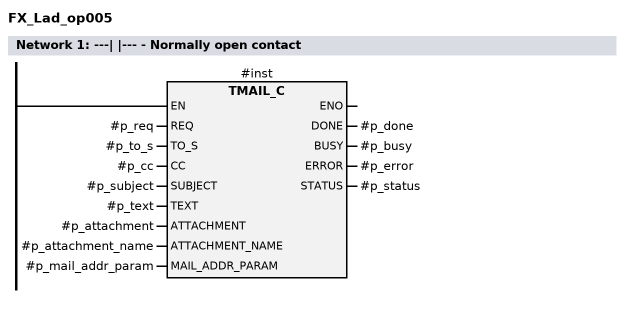
   #inst(REQ := #p_req,   // TMAIL_C
         TO_S := #p_to_s,
         CC := #p_cc,
         SUBJECT := #p_subject,
         TEXT := #p_text,
         ATTACHMENT := #p_attachment,
         ATTACHMENT_NAME := #p_attachment_name,
         MAIL_ADDR_PARAM := #p_mail_addr_param,
         DONE => #p_done,
         BUSY => #p_busy,
         ERROR => #p_error,
         STATUS => #p_status);
END_REGION
END_FUNCTION_BLOCK

FUNCTION_BLOCK "FX_Lad_op021"   // FB349, LAD
{ S7_Optimized_Access := 'TRUE' }
VERSION : 0.1
   VAR_INPUT
      "a" : Bool;
      "b" : Bool;
      c : Bool;
      ia : Int;
      ib : Int;
      ic : Int;
      da : DInt;
      db : DInt;
      ra : Real;
      rb : Real;
      wa : Word;
      wb : Word;
      dwa : DWord;
      ba : Byte;
      ta : Time;
      tb : Time;
      s1 : String;
      s2 : String;
   END_VAR
   VAR_OUTPUT
      q : Bool;
      q2 : Bool;
      io : Int;
      io2 : Int;
      dout : DInt;
      rout : Real;
      wout : Word;
      dwout : DWord;
      bout : Byte;
      tout : Time;
      sout : String;
   END_VAR
   VAR_IN_OUT
      p_req : Bool;
      p_interface : Hw_Interface;
      p_conf_data : Variant;
      p_done : Bool;
      p_busy : Bool;
      p_error : Bool;
      p_status : DWord;
      p_err_loc : DWord;
      arr : Array[0..9] of Int;
      barr : Array[0..7] of Bool;
      iinout : Int;
   END_VAR
   VAR
      inst : T_CONFIG;
      ton1 : TON_TIME;
      tof1 : TOF_TIME;
      tp1 : TP_TIME;
      tonr1 : TONR_TIME;
      ctu1 : CTU_INT;
      ctd1 : CTD_INT;
      ctud1 : CTUD_INT;
      rtrig1 : R_TRIG;
      ftrig1 : F_TRIG;
      edge1 : Bool;
      edge2 : Bool;
      stat1 : Bool;
      stat2 : Bool;
      stati : Int;
   END_VAR
   VAR_TEMP
      t1 : Bool;
      t2 : Bool;
      ti : Int;
      td : DInt;
      tr : Real;
      tw : Word;
      tt : Time;
      var1 : Variant;
   END_VAR
BEGIN

REGION Network 1: ---| |--- - Normally open contact
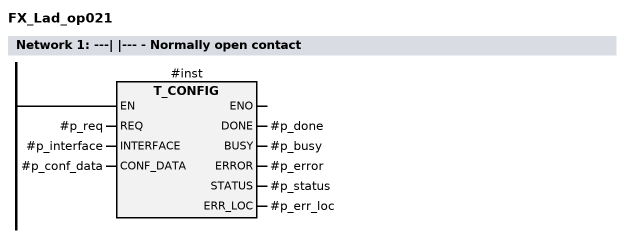
   #inst(Req := #p_req,   // T_CONFIG
         Interface := #p_interface,
         Conf_Data := #p_conf_data,
         Done => #p_done,
         Busy => #p_busy,
         Error => #p_error,
         Status => #p_status,
         Err_Loc => #p_err_loc);
END_REGION
END_FUNCTION_BLOCK

FUNCTION_BLOCK "FB_Lad_Trcv"   // FB350, LAD
{ S7_Optimized_Access := 'TRUE' }
   VAR_INPUT
      en_r : Bool;
      cont : Bool;
      len : UInt;
      id : Conn_Ouc;
      adhoc : Bool;
   END_VAR
   VAR_OUTPUT
      done : Bool;
      busy : Bool;
      err : Bool;
      status : Word;
      rcvdlen : UInt;
   END_VAR
   VAR_IN_OUT
      connect : TCON_IP_v4;
      data : Array[0..99] of Byte;
      comrst : Bool;
      addr : Variant;
   END_VAR
   VAR
      inst : TRCV;
   END_VAR
BEGIN

REGION Network 1: TRCV
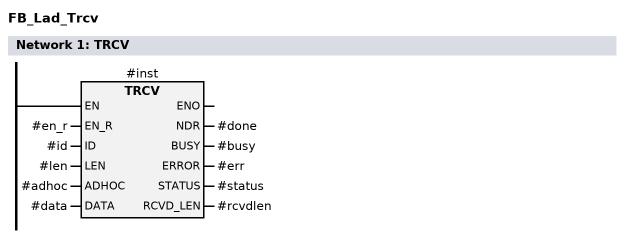
   #inst(EN_R := #en_r,   // TRCV
         ID := #id,
         LEN := #len,
         ADHOC := #adhoc,
         DATA := #data,
         NDR => #done,
         BUSY => #busy,
         ERROR => #err,
         STATUS => #status,
         RCVD_LEN => #rcvdlen);
END_REGION
END_FUNCTION_BLOCK

FUNCTION_BLOCK "FB_Lad_TrcvC"   // FB351, LAD
{ S7_Optimized_Access := 'TRUE' }
   VAR_INPUT
      en_r : Bool;
      cont : Bool;
      len : UInt;
      id : Conn_Ouc;
      adhoc : Bool;
   END_VAR
   VAR_OUTPUT
      done : Bool;
      busy : Bool;
      err : Bool;
      status : Word;
      rcvdlen : UInt;
   END_VAR
   VAR_IN_OUT
      connect : TCON_IP_v4;
      data : Array[0..99] of Byte;
      comrst : Bool;
      addr : Variant;
   END_VAR
   VAR
      inst : TRCV_C;
   END_VAR
BEGIN

REGION Network 1: TRCV_C
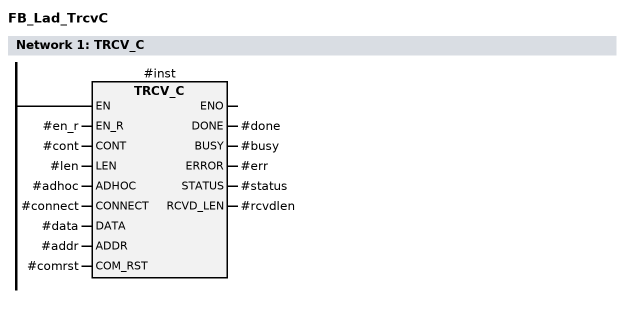
   #inst(EN_R := #en_r,   // TRCV_C
         CONT := #cont,
         LEN := #len,
         ADHOC := #adhoc,
         CONNECT := #connect,
         DATA := #data,
         ADDR := #addr,
         COM_RST := #comrst,
         DONE => #done,
         BUSY => #busy,
         ERROR => #err,
         STATUS => #status,
         RCVD_LEN => #rcvdlen);
END_REGION
END_FUNCTION_BLOCK

FUNCTION_BLOCK "FB_Fbd_TrcvC"   // FB352, FBD
{ S7_Optimized_Access := 'TRUE' }
   VAR_INPUT
      en_r : Bool;
      cont : Bool;
      len : UInt;
      id : Conn_Ouc;
      adhoc : Bool;
   END_VAR
   VAR_OUTPUT
      done : Bool;
      busy : Bool;
      err : Bool;
      status : Word;
      rcvdlen : UInt;
   END_VAR
   VAR_IN_OUT
      connect : TCON_IP_v4;
      data : Array[0..99] of Byte;
      comrst : Bool;
      addr : Variant;
   END_VAR
   VAR
      inst : TRCV_C;
   END_VAR
BEGIN

REGION Network 1: TRCV_C
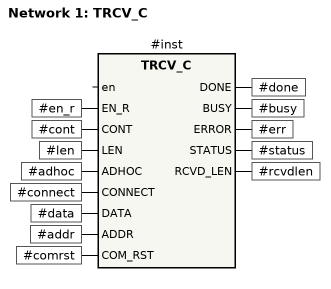
   #inst(EN_R := #en_r,   // TRCV_C
         CONT := #cont,
         LEN := #len,
         ADHOC := #adhoc,
         CONNECT := #connect,
         DATA := #data,
         ADDR := #addr,
         COM_RST := #comrst,
         DONE => #done,
         BUSY => #busy,
         ERROR => #err,
         STATUS => #status,
         RCVD_LEN => #rcvdlen);
END_REGION
END_FUNCTION_BLOCK

FUNCTION_BLOCK "FB_Fbd_Trcv"   // FB353, FBD
{ S7_Optimized_Access := 'TRUE' }
   VAR_INPUT
      en_r : Bool;
      cont : Bool;
      len : UInt;
      id : Conn_Ouc;
      adhoc : Bool;
   END_VAR
   VAR_OUTPUT
      done : Bool;
      busy : Bool;
      err : Bool;
      status : Word;
      rcvdlen : UInt;
   END_VAR
   VAR_IN_OUT
      connect : TCON_IP_v4;
      data : Array[0..99] of Byte;
      comrst : Bool;
      addr : Variant;
   END_VAR
   VAR
      inst : TRCV;
   END_VAR
BEGIN

REGION Network 1: TRCV
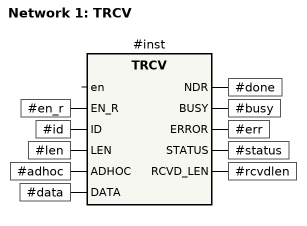
   #inst(EN_R := #en_r,   // TRCV
         ID := #id,
         LEN := #len,
         ADHOC := #adhoc,
         DATA := #data,
         NDR => #done,
         BUSY => #busy,
         ERROR => #err,
         STATUS => #status,
         RCVD_LEN => #rcvdlen);
END_REGION
END_FUNCTION_BLOCK

FUNCTION_BLOCK "FX_Fbd_op005"   // FB354, FBD
{ S7_Optimized_Access := 'TRUE' }
VERSION : 0.1
   VAR_INPUT
      "a" : Bool;
      "b" : Bool;
      c : Bool;
      ia : Int;
      ib : Int;
      ic : Int;
      da : DInt;
      db : DInt;
      ra : Real;
      rb : Real;
      wa : Word;
      wb : Word;
      dwa : DWord;
      ba : Byte;
      ta : Time;
      tb : Time;
      s1 : String;
      s2 : String;
   END_VAR
   VAR_OUTPUT
      q : Bool;
      q2 : Bool;
      io : Int;
      io2 : Int;
      dout : DInt;
      rout : Real;
      wout : Word;
      dwout : DWord;
      bout : Byte;
      tout : Time;
      sout : String;
   END_VAR
   VAR_IN_OUT
      p_req : Bool;
      p_to_s : String;
      p_cc : String;
      p_subject : String;
      p_text : String;
      p_attachment : Variant;
      p_attachment_name : String;
      p_mail_addr_param : Variant;
      p_done : Bool;
      p_busy : Bool;
      p_error : Bool;
      p_status : Word;
      arr : Array[0..9] of Int;
      barr : Array[0..7] of Bool;
      iinout : Int;
   END_VAR
   VAR
      inst : TMAIL_C;
      ton1 : TON_TIME;
      tof1 : TOF_TIME;
      tp1 : TP_TIME;
      tonr1 : TONR_TIME;
      ctu1 : CTU_INT;
      ctd1 : CTD_INT;
      ctud1 : CTUD_INT;
      rtrig1 : R_TRIG;
      ftrig1 : F_TRIG;
      edge1 : Bool;
      edge2 : Bool;
      stat1 : Bool;
      stat2 : Bool;
      stati : Int;
   END_VAR
   VAR_TEMP
      t1 : Bool;
      t2 : Bool;
      ti : Int;
      td : DInt;
      tr : Real;
      tw : Word;
      tt : Time;
      var1 : Variant;
   END_VAR
BEGIN

REGION Network 1: ---| |--- - Normally open contact
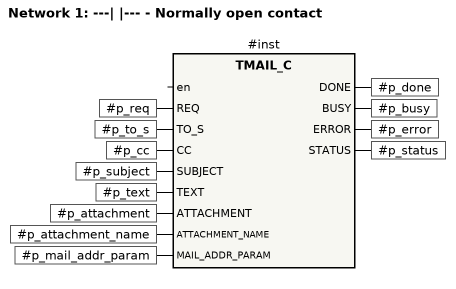
   #inst(REQ := #p_req,   // TMAIL_C
         TO_S := #p_to_s,
         CC := #p_cc,
         SUBJECT := #p_subject,
         TEXT := #p_text,
         ATTACHMENT := #p_attachment,
         ATTACHMENT_NAME := #p_attachment_name,
         MAIL_ADDR_PARAM := #p_mail_addr_param,
         DONE => #p_done,
         BUSY => #p_busy,
         ERROR => #p_error,
         STATUS => #p_status);
END_REGION
END_FUNCTION_BLOCK

FUNCTION_BLOCK "FX_Fbd_op021"   // FB355, FBD
{ S7_Optimized_Access := 'TRUE' }
VERSION : 0.1
   VAR_INPUT
      "a" : Bool;
      "b" : Bool;
      c : Bool;
      ia : Int;
      ib : Int;
      ic : Int;
      da : DInt;
      db : DInt;
      ra : Real;
      rb : Real;
      wa : Word;
      wb : Word;
      dwa : DWord;
      ba : Byte;
      ta : Time;
      tb : Time;
      s1 : String;
      s2 : String;
   END_VAR
   VAR_OUTPUT
      q : Bool;
      q2 : Bool;
      io : Int;
      io2 : Int;
      dout : DInt;
      rout : Real;
      wout : Word;
      dwout : DWord;
      bout : Byte;
      tout : Time;
      sout : String;
   END_VAR
   VAR_IN_OUT
      p_req : Bool;
      p_interface : Hw_Interface;
      p_conf_data : Variant;
      p_done : Bool;
      p_busy : Bool;
      p_error : Bool;
      p_status : DWord;
      p_err_loc : DWord;
      arr : Array[0..9] of Int;
      barr : Array[0..7] of Bool;
      iinout : Int;
   END_VAR
   VAR
      inst : T_CONFIG;
      ton1 : TON_TIME;
      tof1 : TOF_TIME;
      tp1 : TP_TIME;
      tonr1 : TONR_TIME;
      ctu1 : CTU_INT;
      ctd1 : CTD_INT;
      ctud1 : CTUD_INT;
      rtrig1 : R_TRIG;
      ftrig1 : F_TRIG;
      edge1 : Bool;
      edge2 : Bool;
      stat1 : Bool;
      stat2 : Bool;
      stati : Int;
   END_VAR
   VAR_TEMP
      t1 : Bool;
      t2 : Bool;
      ti : Int;
      td : DInt;
      tr : Real;
      tw : Word;
      tt : Time;
      var1 : Variant;
   END_VAR
BEGIN

REGION Network 1: ---| |--- - Normally open contact
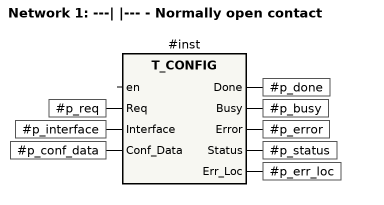
   #inst(Req := #p_req,   // T_CONFIG
         Interface := #p_interface,
         Conf_Data := #p_conf_data,
         Done => #p_done,
         Busy => #p_busy,
         Error => #p_error,
         Status => #p_status,
         Err_Loc => #p_err_loc);
END_REGION
END_FUNCTION_BLOCK

FUNCTION_BLOCK "FB_Lad_ex051"   // FB356, LAD
{ S7_Optimized_Access := 'TRUE' }
   VAR_INPUT
      v_mode : Int;
      v_f_id : Hw_Io;
      v_mlen : UInt;
   END_VAR
   VAR_OUTPUT
      v_new : Bool;
      v_status : DWord;
      v_id : Hw_Io;
      v_len : UInt;
   END_VAR
   VAR_IN_OUT
      v_tinfo : Array[0..99] of Byte;
      v_ainfo : Array[0..99] of Byte;
   END_VAR
   VAR
      inst : RALRM;
   END_VAR
BEGIN

REGION Network 1: Description RALRM
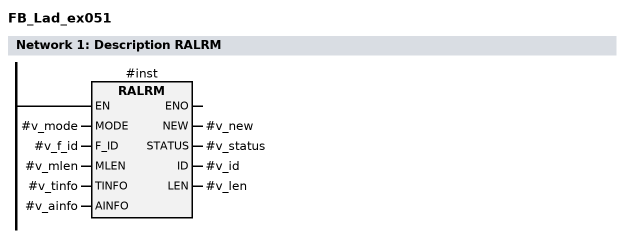
   #inst(MODE := #v_mode,   // RALRM
         F_ID := #v_f_id,
         MLEN := #v_mlen,
         TINFO := #v_tinfo,
         AINFO := #v_ainfo,
         NEW => #v_new,
         STATUS => #v_status,
         ID => #v_id,
         LEN => #v_len);
END_REGION
END_FUNCTION_BLOCK

FUNCTION_BLOCK "FB_Lad_ex071"   // FB357, LAD
{ S7_Optimized_Access := 'TRUE' }
   VAR_INPUT
      v_com_rst : Bool;
      v_start : Bool;
      v_end : Bool;
   END_VAR
   VAR_OUTPUT
      v_status : DWord;
   END_VAR
   VAR_IN_OUT
      v_penergy : PE_PLUS;
   END_VAR
   VAR
      inst : PE_WOL;
   END_VAR
BEGIN

REGION Network 1: Description PE_WOL
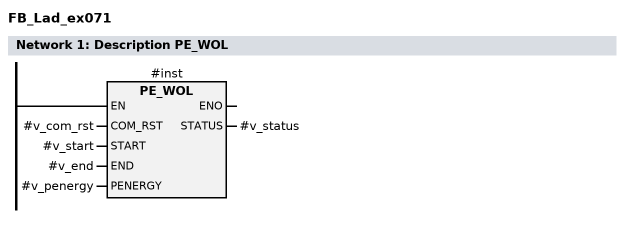
   #inst(COM_RST := #v_com_rst, START := #v_start, END := #v_end, PENERGY := #v_penergy, STATUS => #v_status);   // PE_WOL
END_REGION
END_FUNCTION_BLOCK

FUNCTION_BLOCK "FX_Lad_ex037"   // FB358, LAD
{ S7_Optimized_Access := 'TRUE' }
VERSION : 0.1
   VAR_INPUT
      "a" : Bool;
      "b" : Bool;
      c : Bool;
      ia : Int;
      ib : Int;
      ic : Int;
      da : DInt;
      db : DInt;
      ra : Real;
      rb : Real;
      wa : Word;
      wb : Word;
      dwa : DWord;
      ba : Byte;
      ta : Time;
      tb : Time;
      s1 : String;
      s2 : String;
   END_VAR
   VAR_OUTPUT
      q : Bool;
      q2 : Bool;
      io : Int;
      io2 : Int;
      dout : DInt;
      rout : Real;
      wout : Word;
      dwout : DWord;
      bout : Byte;
      tout : Time;
      sout : String;
   END_VAR
   VAR_IN_OUT
      x_wstring : WString;
      arr : Array[0..9] of Int;
      barr : Array[0..7] of Bool;
      iinout : Int;
   END_VAR
   VAR
      ton1 : TON_TIME;
      tof1 : TOF_TIME;
      tp1 : TP_TIME;
      tonr1 : TONR_TIME;
      ctu1 : CTU_INT;
      ctd1 : CTD_INT;
      ctud1 : CTUD_INT;
      rtrig1 : R_TRIG;
      ftrig1 : F_TRIG;
      edge1 : Bool;
      edge2 : Bool;
      stat1 : Bool;
      stat2 : Bool;
      stati : Int;
   END_VAR
   VAR_TEMP
      t1 : Bool;
      t2 : Bool;
      ti : Int;
      td : DInt;
      tr : Real;
      tw : Word;
      tt : Time;
      var1 : Variant;
   END_VAR
BEGIN

REGION Network 1: ---| |--- - Normally open contact
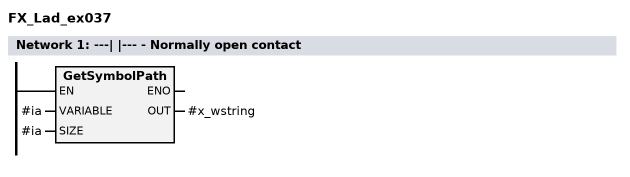
   // no SCL statement known for GetSymbolPath: written as a call
   #x_wstring := GetSymbolPath(variable := #ia, size := #ia);
END_REGION
END_FUNCTION_BLOCK

FUNCTION_BLOCK "FX_Lad_ex051"   // FB359, LAD
{ S7_Optimized_Access := 'TRUE' }
VERSION : 0.1
   VAR_INPUT
      "a" : Bool;
      "b" : Bool;
      c : Bool;
      ia : Int;
      ib : Int;
      ic : Int;
      da : DInt;
      db : DInt;
      ra : Real;
      rb : Real;
      wa : Word;
      wb : Word;
      dwa : DWord;
      ba : Byte;
      ta : Time;
      tb : Time;
      s1 : String;
      s2 : String;
   END_VAR
   VAR_OUTPUT
      q : Bool;
      q2 : Bool;
      io : Int;
      io2 : Int;
      dout : DInt;
      rout : Real;
      wout : Word;
      dwout : DWord;
      bout : Byte;
      tout : Time;
      sout : String;
   END_VAR
   VAR_IN_OUT
      p_mode : Int;
      p_f_id : Hw_Io;
      p_mlen : UInt;
      p_new : Bool;
      p_status : DWord;
      p_id : Hw_Io;
      p_len : UInt;
      p_tinfo : Variant;
      p_ainfo : Variant;
      arr : Array[0..9] of Int;
      barr : Array[0..7] of Bool;
      iinout : Int;
   END_VAR
   VAR
      inst : RALRM;
      ton1 : TON_TIME;
      tof1 : TOF_TIME;
      tp1 : TP_TIME;
      tonr1 : TONR_TIME;
      ctu1 : CTU_INT;
      ctd1 : CTD_INT;
      ctud1 : CTUD_INT;
      rtrig1 : R_TRIG;
      ftrig1 : F_TRIG;
      edge1 : Bool;
      edge2 : Bool;
      stat1 : Bool;
      stat2 : Bool;
      stati : Int;
   END_VAR
   VAR_TEMP
      t1 : Bool;
      t2 : Bool;
      ti : Int;
      td : DInt;
      tr : Real;
      tw : Word;
      tt : Time;
      var1 : Variant;
   END_VAR
BEGIN

REGION Network 1: ---| |--- - Normally open contact
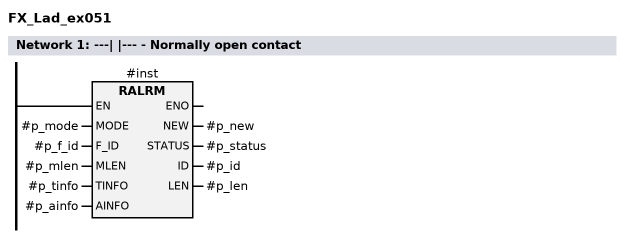
   #inst(MODE := #p_mode,   // RALRM
         F_ID := #p_f_id,
         MLEN := #p_mlen,
         TINFO := #p_tinfo,
         AINFO := #p_ainfo,
         NEW => #p_new,
         STATUS => #p_status,
         ID => #p_id,
         LEN => #p_len);
END_REGION
END_FUNCTION_BLOCK

FUNCTION_BLOCK "FB_Fbd_ex037"   // FB360, FBD
{ S7_Optimized_Access := 'TRUE' }
   VAR_INPUT
      v_size : DInt;
   END_VAR
   VAR_OUTPUT
      v_out : WString;
   END_VAR
   VAR_IN_OUT
      v_variable : Variant;
   END_VAR
BEGIN

REGION Network 1: Querying GetSymbolPath - actual parameter at beginning of a call path
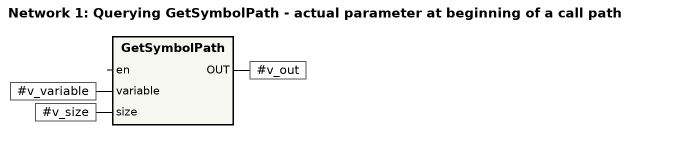
   // no SCL statement known for GetSymbolPath: written as a call
   #v_out := GetSymbolPath(variable := #v_variable, size := #v_size);
END_REGION
END_FUNCTION_BLOCK

FUNCTION_BLOCK "FB_Fbd_ex051"   // FB361, FBD
{ S7_Optimized_Access := 'TRUE' }
   VAR_INPUT
      v_mode : Int;
      v_f_id : Hw_Io;
      v_mlen : UInt;
   END_VAR
   VAR_OUTPUT
      v_new : Bool;
      v_status : DWord;
      v_id : Hw_Io;
      v_len : UInt;
   END_VAR
   VAR_IN_OUT
      v_tinfo : Array[0..99] of Byte;
      v_ainfo : Array[0..99] of Byte;
   END_VAR
   VAR
      inst : RALRM;
   END_VAR
BEGIN

REGION Network 1: Description RALRM
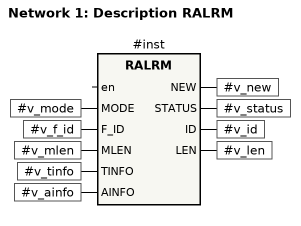
   #inst(MODE := #v_mode,   // RALRM
         F_ID := #v_f_id,
         MLEN := #v_mlen,
         TINFO := #v_tinfo,
         AINFO := #v_ainfo,
         NEW => #v_new,
         STATUS => #v_status,
         ID => #v_id,
         LEN => #v_len);
END_REGION
END_FUNCTION_BLOCK

FUNCTION_BLOCK "FB_Fbd_ex071"   // FB362, FBD
{ S7_Optimized_Access := 'TRUE' }
   VAR_INPUT
      v_com_rst : Bool;
      v_start : Bool;
      v_end : Bool;
   END_VAR
   VAR_OUTPUT
      v_status : DWord;
   END_VAR
   VAR_IN_OUT
      v_penergy : PE_PLUS;
   END_VAR
   VAR
      inst : PE_WOL;
   END_VAR
BEGIN

REGION Network 1: Description PE_WOL
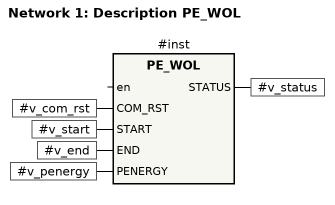
   #inst(COM_RST := #v_com_rst, START := #v_start, END := #v_end, PENERGY := #v_penergy, STATUS => #v_status);   // PE_WOL
END_REGION
END_FUNCTION_BLOCK

FUNCTION_BLOCK "FX_Lad_095"   // FB363, LAD
{ S7_Optimized_Access := 'TRUE' }
VERSION : 0.1
   VAR_INPUT
      "a" : Bool;
      "b" : Bool;
      c : Bool;
      ia : Int;
      ib : Int;
      ic : Int;
      da : DInt;
      db : DInt;
      ra : Real;
      rb : Real;
      wa : Word;
      wb : Word;
      dwa : DWord;
      ba : Byte;
      ta : Time;
      tb : Time;
      s1 : String;
      s2 : String;
   END_VAR
   VAR_OUTPUT
      q : Bool;
      q2 : Bool;
      io : Int;
      io2 : Int;
      dout : DInt;
      rout : Real;
      wout : Word;
      dwout : DWord;
      bout : Byte;
      tout : Time;
      sout : String;
   END_VAR
   VAR_IN_OUT
      x_usint : USInt;
      arr : Array[0..9] of Int;
      barr : Array[0..7] of Bool;
      iinout : Int;
   END_VAR
   VAR
      ton1 : TON_TIME;
      tof1 : TOF_TIME;
      tp1 : TP_TIME;
      tonr1 : TONR_TIME;
      ctu1 : CTU_INT;
      ctd1 : CTD_INT;
      ctud1 : CTUD_INT;
      rtrig1 : R_TRIG;
      ftrig1 : F_TRIG;
      edge1 : Bool;
      edge2 : Bool;
      stat1 : Bool;
      stat2 : Bool;
      stati : Int;
   END_VAR
   VAR_TEMP
      t1 : Bool;
      t2 : Bool;
      ti : Int;
      td : DInt;
      tr : Real;
      tw : Word;
      tt : Time;
      var1 : Variant;
   END_VAR
BEGIN

REGION Network 1: ---| |--- - Normally open contact
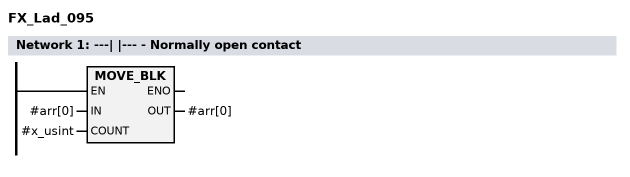
   MOVE_BLK(IN := #arr[0], COUNT := #x_usint, OUT => #arr[0]);
END_REGION
END_FUNCTION_BLOCK

FUNCTION_BLOCK "FX_Lad_097"   // FB364, LAD
{ S7_Optimized_Access := 'TRUE' }
VERSION : 0.1
   VAR_INPUT
      "a" : Bool;
      "b" : Bool;
      c : Bool;
      ia : Int;
      ib : Int;
      ic : Int;
      da : DInt;
      db : DInt;
      ra : Real;
      rb : Real;
      wa : Word;
      wb : Word;
      dwa : DWord;
      ba : Byte;
      ta : Time;
      tb : Time;
      s1 : String;
      s2 : String;
   END_VAR
   VAR_OUTPUT
      q : Bool;
      q2 : Bool;
      io : Int;
      io2 : Int;
      dout : DInt;
      rout : Real;
      wout : Word;
      dwout : DWord;
      bout : Byte;
      tout : Time;
      sout : String;
   END_VAR
   VAR_IN_OUT
      x_usint : USInt;
      arr : Array[0..9] of Int;
      barr : Array[0..7] of Bool;
      iinout : Int;
   END_VAR
   VAR
      ton1 : TON_TIME;
      tof1 : TOF_TIME;
      tp1 : TP_TIME;
      tonr1 : TONR_TIME;
      ctu1 : CTU_INT;
      ctd1 : CTD_INT;
      ctud1 : CTUD_INT;
      rtrig1 : R_TRIG;
      ftrig1 : F_TRIG;
      edge1 : Bool;
      edge2 : Bool;
      stat1 : Bool;
      stat2 : Bool;
      stati : Int;
   END_VAR
   VAR_TEMP
      t1 : Bool;
      t2 : Bool;
      ti : Int;
      td : DInt;
      tr : Real;
      tw : Word;
      tt : Time;
      var1 : Variant;
   END_VAR
BEGIN

REGION Network 1: ---| |--- - Normally open contact
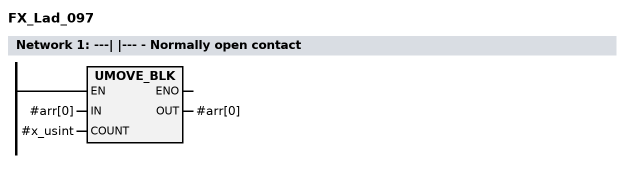
   UMOVE_BLK(IN := #arr[0], COUNT := #x_usint, OUT => #arr[0]);
END_REGION
END_FUNCTION_BLOCK

FUNCTION_BLOCK "FX_Lad_098"   // FB365, LAD
{ S7_Optimized_Access := 'TRUE' }
VERSION : 0.1
   VAR_INPUT
      "a" : Bool;
      "b" : Bool;
      c : Bool;
      ia : Int;
      ib : Int;
      ic : Int;
      da : DInt;
      db : DInt;
      ra : Real;
      rb : Real;
      wa : Word;
      wb : Word;
      dwa : DWord;
      ba : Byte;
      ta : Time;
      tb : Time;
      s1 : String;
      s2 : String;
   END_VAR
   VAR_OUTPUT
      q : Bool;
      q2 : Bool;
      io : Int;
      io2 : Int;
      dout : DInt;
      rout : Real;
      wout : Word;
      dwout : DWord;
      bout : Byte;
      tout : Time;
      sout : String;
   END_VAR
   VAR_IN_OUT
      p_in : Date;
      p_count : USInt;
      p_out : Date;
      s_in : Int;
      s_count : UDInt;
      s_out : Array[0..9] of Int;
      arr : Array[0..9] of Int;
      barr : Array[0..7] of Bool;
      iinout : Int;
   END_VAR
   VAR
      ton1 : TON_TIME;
      tof1 : TOF_TIME;
      tp1 : TP_TIME;
      tonr1 : TONR_TIME;
      ctu1 : CTU_INT;
      ctd1 : CTD_INT;
      ctud1 : CTUD_INT;
      rtrig1 : R_TRIG;
      ftrig1 : F_TRIG;
      edge1 : Bool;
      edge2 : Bool;
      stat1 : Bool;
      stat2 : Bool;
      stati : Int;
   END_VAR
   VAR_TEMP
      t1 : Bool;
      t2 : Bool;
      ti : Int;
      td : DInt;
      tr : Real;
      tw : Word;
      tt : Time;
      var1 : Variant;
   END_VAR
BEGIN

REGION Network 1: ---| |--- - Normally open contact
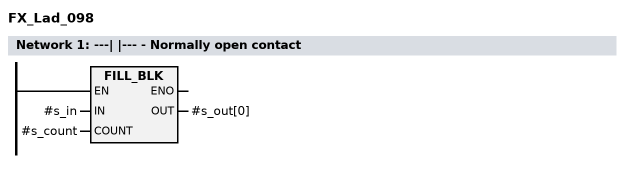
   RUNG wire#powerrail
      FillBlockI(in := #s_in, count := #s_count, out => #s_out[0])
   END_RUNG
   // the same network as SCL:
   FILL_BLK(IN := #s_in, COUNT := #s_count, OUT => #s_out[0]);
END_REGION
END_FUNCTION_BLOCK

FUNCTION_BLOCK "FX_Lad_099"   // FB366, LAD
{ S7_Optimized_Access := 'TRUE' }
VERSION : 0.1
   VAR_INPUT
      "a" : Bool;
      "b" : Bool;
      c : Bool;
      ia : Int;
      ib : Int;
      ic : Int;
      da : DInt;
      db : DInt;
      ra : Real;
      rb : Real;
      wa : Word;
      wb : Word;
      dwa : DWord;
      ba : Byte;
      ta : Time;
      tb : Time;
      s1 : String;
      s2 : String;
   END_VAR
   VAR_OUTPUT
      q : Bool;
      q2 : Bool;
      io : Int;
      io2 : Int;
      dout : DInt;
      rout : Real;
      wout : Word;
      dwout : DWord;
      bout : Byte;
      tout : Time;
      sout : String;
   END_VAR
   VAR_IN_OUT
      p_in : Date;
      p_count : USInt;
      p_out : Date;
      s_in : Int;
      s_count : UDInt;
      s_out : Array[0..9] of Int;
      arr : Array[0..9] of Int;
      barr : Array[0..7] of Bool;
      iinout : Int;
   END_VAR
   VAR
      ton1 : TON_TIME;
      tof1 : TOF_TIME;
      tp1 : TP_TIME;
      tonr1 : TONR_TIME;
      ctu1 : CTU_INT;
      ctd1 : CTD_INT;
      ctud1 : CTUD_INT;
      rtrig1 : R_TRIG;
      ftrig1 : F_TRIG;
      edge1 : Bool;
      edge2 : Bool;
      stat1 : Bool;
      stat2 : Bool;
      stati : Int;
   END_VAR
   VAR_TEMP
      t1 : Bool;
      t2 : Bool;
      ti : Int;
      td : DInt;
      tr : Real;
      tw : Word;
      tt : Time;
      var1 : Variant;
   END_VAR
BEGIN

REGION Network 1: ---| |--- - Normally open contact
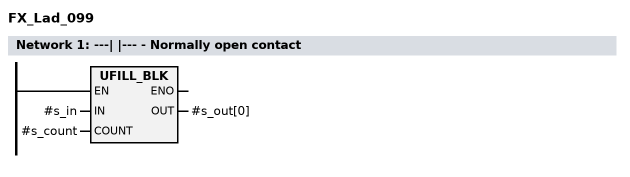
   UFILL_BLK(IN := #s_in, COUNT := #s_count, OUT => #s_out[0]);
END_REGION
END_FUNCTION_BLOCK

FUNCTION_BLOCK "FX_Fbd_100"   // FB367, FBD
{ S7_Optimized_Access := 'TRUE' }
VERSION : 0.1
   VAR_INPUT
      "a" : Bool;
      "b" : Bool;
      c : Bool;
      ia : Int;
      ib : Int;
      ic : Int;
      da : DInt;
      db : DInt;
      ra : Real;
      rb : Real;
      wa : Word;
      wb : Word;
      dwa : DWord;
      ba : Byte;
      ta : Time;
      tb : Time;
      s1 : String;
      s2 : String;
   END_VAR
   VAR_OUTPUT
      q : Bool;
      q2 : Bool;
      io : Int;
      io2 : Int;
      dout : DInt;
      rout : Real;
      wout : Word;
      dwout : DWord;
      bout : Byte;
      tout : Time;
      sout : String;
   END_VAR
   VAR_IN_OUT
      x_usint : USInt;
      arr : Array[0..9] of Int;
      barr : Array[0..7] of Bool;
      iinout : Int;
   END_VAR
   VAR
      ton1 : TON_TIME;
      tof1 : TOF_TIME;
      tp1 : TP_TIME;
      tonr1 : TONR_TIME;
      ctu1 : CTU_INT;
      ctd1 : CTD_INT;
      ctud1 : CTUD_INT;
      rtrig1 : R_TRIG;
      ftrig1 : F_TRIG;
      edge1 : Bool;
      edge2 : Bool;
      stat1 : Bool;
      stat2 : Bool;
      stati : Int;
   END_VAR
   VAR_TEMP
      t1 : Bool;
      t2 : Bool;
      ti : Int;
      td : DInt;
      tr : Real;
      tw : Word;
      tt : Time;
      var1 : Variant;
   END_VAR
BEGIN

REGION Network 1: ---| |--- - Normally open contact
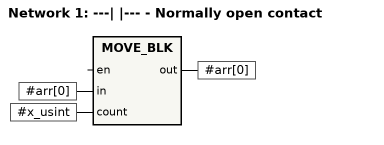
   MOVE_BLK(IN := #arr[0], COUNT := #x_usint, OUT => #arr[0]);
END_REGION
END_FUNCTION_BLOCK

FUNCTION_BLOCK "FX_Fbd_102"   // FB368, FBD
{ S7_Optimized_Access := 'TRUE' }
VERSION : 0.1
   VAR_INPUT
      "a" : Bool;
      "b" : Bool;
      c : Bool;
      ia : Int;
      ib : Int;
      ic : Int;
      da : DInt;
      db : DInt;
      ra : Real;
      rb : Real;
      wa : Word;
      wb : Word;
      dwa : DWord;
      ba : Byte;
      ta : Time;
      tb : Time;
      s1 : String;
      s2 : String;
   END_VAR
   VAR_OUTPUT
      q : Bool;
      q2 : Bool;
      io : Int;
      io2 : Int;
      dout : DInt;
      rout : Real;
      wout : Word;
      dwout : DWord;
      bout : Byte;
      tout : Time;
      sout : String;
   END_VAR
   VAR_IN_OUT
      x_usint : USInt;
      arr : Array[0..9] of Int;
      barr : Array[0..7] of Bool;
      iinout : Int;
   END_VAR
   VAR
      ton1 : TON_TIME;
      tof1 : TOF_TIME;
      tp1 : TP_TIME;
      tonr1 : TONR_TIME;
      ctu1 : CTU_INT;
      ctd1 : CTD_INT;
      ctud1 : CTUD_INT;
      rtrig1 : R_TRIG;
      ftrig1 : F_TRIG;
      edge1 : Bool;
      edge2 : Bool;
      stat1 : Bool;
      stat2 : Bool;
      stati : Int;
   END_VAR
   VAR_TEMP
      t1 : Bool;
      t2 : Bool;
      ti : Int;
      td : DInt;
      tr : Real;
      tw : Word;
      tt : Time;
      var1 : Variant;
   END_VAR
BEGIN

REGION Network 1: ---| |--- - Normally open contact
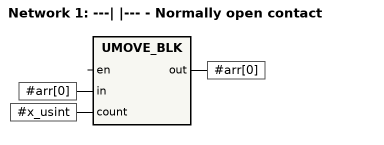
   UMOVE_BLK(IN := #arr[0], COUNT := #x_usint, OUT => #arr[0]);
END_REGION
END_FUNCTION_BLOCK

FUNCTION_BLOCK "FX_Fbd_103"   // FB369, FBD
{ S7_Optimized_Access := 'TRUE' }
VERSION : 0.1
   VAR_INPUT
      "a" : Bool;
      "b" : Bool;
      c : Bool;
      ia : Int;
      ib : Int;
      ic : Int;
      da : DInt;
      db : DInt;
      ra : Real;
      rb : Real;
      wa : Word;
      wb : Word;
      dwa : DWord;
      ba : Byte;
      ta : Time;
      tb : Time;
      s1 : String;
      s2 : String;
   END_VAR
   VAR_OUTPUT
      q : Bool;
      q2 : Bool;
      io : Int;
      io2 : Int;
      dout : DInt;
      rout : Real;
      wout : Word;
      dwout : DWord;
      bout : Byte;
      tout : Time;
      sout : String;
   END_VAR
   VAR_IN_OUT
      p_in : Date;
      p_count : USInt;
      p_out : Date;
      s_in : Int;
      s_count : UDInt;
      s_out : Array[0..9] of Int;
      arr : Array[0..9] of Int;
      barr : Array[0..7] of Bool;
      iinout : Int;
   END_VAR
   VAR
      ton1 : TON_TIME;
      tof1 : TOF_TIME;
      tp1 : TP_TIME;
      tonr1 : TONR_TIME;
      ctu1 : CTU_INT;
      ctd1 : CTD_INT;
      ctud1 : CTUD_INT;
      rtrig1 : R_TRIG;
      ftrig1 : F_TRIG;
      edge1 : Bool;
      edge2 : Bool;
      stat1 : Bool;
      stat2 : Bool;
      stati : Int;
   END_VAR
   VAR_TEMP
      t1 : Bool;
      t2 : Bool;
      ti : Int;
      td : DInt;
      tr : Real;
      tw : Word;
      tt : Time;
      var1 : Variant;
   END_VAR
BEGIN

REGION Network 1: ---| |--- - Normally open contact
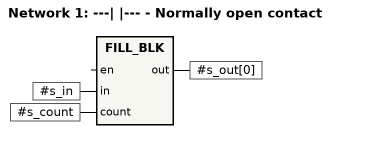
   FILL_BLK(IN := #s_in, COUNT := #s_count, OUT => #s_out[0]);
END_REGION
END_FUNCTION_BLOCK

FUNCTION_BLOCK "FX_Fbd_104"   // FB370, FBD
{ S7_Optimized_Access := 'TRUE' }
VERSION : 0.1
   VAR_INPUT
      "a" : Bool;
      "b" : Bool;
      c : Bool;
      ia : Int;
      ib : Int;
      ic : Int;
      da : DInt;
      db : DInt;
      ra : Real;
      rb : Real;
      wa : Word;
      wb : Word;
      dwa : DWord;
      ba : Byte;
      ta : Time;
      tb : Time;
      s1 : String;
      s2 : String;
   END_VAR
   VAR_OUTPUT
      q : Bool;
      q2 : Bool;
      io : Int;
      io2 : Int;
      dout : DInt;
      rout : Real;
      wout : Word;
      dwout : DWord;
      bout : Byte;
      tout : Time;
      sout : String;
   END_VAR
   VAR_IN_OUT
      p_in : Date;
      p_count : USInt;
      p_out : Date;
      s_in : Int;
      s_count : UDInt;
      s_out : Array[0..9] of Int;
      arr : Array[0..9] of Int;
      barr : Array[0..7] of Bool;
      iinout : Int;
   END_VAR
   VAR
      ton1 : TON_TIME;
      tof1 : TOF_TIME;
      tp1 : TP_TIME;
      tonr1 : TONR_TIME;
      ctu1 : CTU_INT;
      ctd1 : CTD_INT;
      ctud1 : CTUD_INT;
      rtrig1 : R_TRIG;
      ftrig1 : F_TRIG;
      edge1 : Bool;
      edge2 : Bool;
      stat1 : Bool;
      stat2 : Bool;
      stati : Int;
   END_VAR
   VAR_TEMP
      t1 : Bool;
      t2 : Bool;
      ti : Int;
      td : DInt;
      tr : Real;
      tw : Word;
      tt : Time;
      var1 : Variant;
   END_VAR
BEGIN

REGION Network 1: ---| |--- - Normally open contact
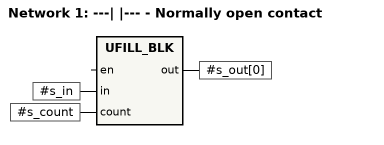
   UFILL_BLK(IN := #s_in, COUNT := #s_count, OUT => #s_out[0]);
END_REGION
END_FUNCTION_BLOCK

FUNCTION_BLOCK "FX_Lad_ex001"   // FB371, LAD
{ S7_Optimized_Access := 'TRUE' }
VERSION : 0.1
   VAR_INPUT
      "a" : Bool;
      "b" : Bool;
      c : Bool;
      ia : Int;
      ib : Int;
      ic : Int;
      da : DInt;
      db : DInt;
      ra : Real;
      rb : Real;
      wa : Word;
      wb : Word;
      dwa : DWord;
      ba : Byte;
      ta : Time;
      tb : Time;
      s1 : String;
      s2 : String;
   END_VAR
   VAR_OUTPUT
      q : Bool;
      q2 : Bool;
      io : Int;
      io2 : Int;
      dout : DInt;
      rout : Real;
      wout : Word;
      dwout : DWord;
      bout : Byte;
      tout : Time;
      sout : String;
   END_VAR
   VAR_IN_OUT
      p0 : DTL;
      p1 : DTL;
      arr : Array[0..9] of Int;
      barr : Array[0..7] of Bool;
      iinout : Int;
   END_VAR
   VAR
      ton1 : TON_TIME;
      tof1 : TOF_TIME;
      tp1 : TP_TIME;
      tonr1 : TONR_TIME;
      ctu1 : CTU_INT;
      ctd1 : CTD_INT;
      ctud1 : CTUD_INT;
      rtrig1 : R_TRIG;
      ftrig1 : F_TRIG;
      edge1 : Bool;
      edge2 : Bool;
      stat1 : Bool;
      stat2 : Bool;
      stati : Int;
   END_VAR
   VAR_TEMP
      t1 : Bool;
      t2 : Bool;
      ti : Int;
      td : DInt;
      tr : Real;
      tw : Word;
      tt : Time;
      var1 : Variant;
   END_VAR
BEGIN

REGION Network 1: ---| |--- - Normally open contact
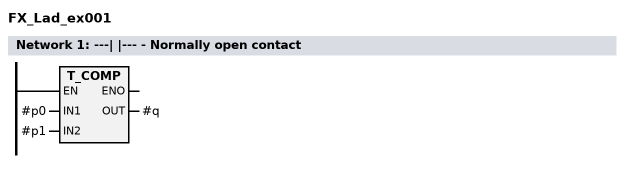
   T_COMP(IN1 := #p0, IN2 := #p1, OUT => #q);
END_REGION
END_FUNCTION_BLOCK

FUNCTION_BLOCK "FX_Lad_ex016"   // FB372, LAD
{ S7_Optimized_Access := 'TRUE' }
VERSION : 0.1
   VAR_INPUT
      "a" : Bool;
      "b" : Bool;
      c : Bool;
      ia : Int;
      ib : Int;
      ic : Int;
      da : DInt;
      db : DInt;
      ra : Real;
      rb : Real;
      wa : Word;
      wb : Word;
      dwa : DWord;
      ba : Byte;
      ta : Time;
      tb : Time;
      s1 : String;
      s2 : String;
   END_VAR
   VAR_OUTPUT
      q : Bool;
      q2 : Bool;
      io : Int;
      io2 : Int;
      dout : DInt;
      rout : Real;
      wout : Word;
      dwout : DWord;
      bout : Byte;
      tout : Time;
      sout : String;
   END_VAR
   VAR_IN_OUT
      p0 : String;
      p1 : String;
      arr : Array[0..9] of Int;
      barr : Array[0..7] of Bool;
      iinout : Int;
   END_VAR
   VAR
      ton1 : TON_TIME;
      tof1 : TOF_TIME;
      tp1 : TP_TIME;
      tonr1 : TONR_TIME;
      ctu1 : CTU_INT;
      ctd1 : CTD_INT;
      ctud1 : CTUD_INT;
      rtrig1 : R_TRIG;
      ftrig1 : F_TRIG;
      edge1 : Bool;
      edge2 : Bool;
      stat1 : Bool;
      stat2 : Bool;
      stati : Int;
   END_VAR
   VAR_TEMP
      t1 : Bool;
      t2 : Bool;
      ti : Int;
      td : DInt;
      tr : Real;
      tw : Word;
      tt : Time;
      var1 : Variant;
   END_VAR
BEGIN

REGION Network 1: ---| |--- - Normally open contact
